(*
SPDX-FileCopyrightText: © 2026 Oleksandr Tiutyk <trofimich@gmail.com>
SPDX-License-Identifier: MIT
License: https://opensource.org/license/mit
*)

(*!
<summary>
Beckhoff EP1008_0001: 8-channel digital input EtherCAT Box (24 V DC, 3 ms filter, M8).
</summary>
<description>
Process image mapping structure for the EP1008_0001 EtherCAT Box IP67 module with 8 discrete inputs.
When used for I/O, link located fields or their containing buffers to the matching selected PDOs.
The record is not a packed wire buffer; compiler padding is not part of the device specification.
Unlinked/default values do not prove valid I/O. The caller evaluates bus/channel validity before use.
Use one owner task per instance and externally synchronize other access; multi-field snapshots are not atomic.
Copies store data without creating hardware links. Keep borrowed field references valid while consumers are bound.
This passive record performs no validation, synchronization, configuration or protocol advancement.
</description>
*)
TYPE EP1008_0001 :
STRUCT
	Ch1 AT %I* : BOOL;
	Ch2 AT %I* : BOOL;
	Ch3 AT %I* : BOOL;
	Ch4 AT %I* : BOOL;
	Ch5 AT %I* : BOOL;
	Ch6 AT %I* : BOOL;
	Ch7 AT %I* : BOOL;
	Ch8 AT %I* : BOOL;
END_STRUCT
END_TYPE

(* stored: Version 1.1.0.1, ProductVersion 3.1.4026.20
   DUT EP1008_0001: Id {b12a82c4-163f-496c-90a1-f54772aa7671} *)
